// TIA Portal V20 export
FUNCTION_BLOCK "FB_Motor"   // FB102, LAD
TITLE = Direct-on-line motor with running feedback and trip monitoring
{ S7_Optimized_Access := 'TRUE' }
AUTHOR : Demo
VERSION : 0.2
// LAD version. Same interface as scl/14_FB_Motor.scl.
// stored: AutoNumber false, SetENOAutomatically false
   VAR_INPUT
      Run : Bool;   // Request: run the motor
      Permit : Bool := true;   // Interlock: motor may only run when TRUE
      RunFb : Bool;   // Running feedback (contactor auxiliary contact)
      Trip : Bool;   // Motor protection breaker tripped
      FeedbackTime : Time := T#5S;   // Max time from command to feedback
   END_VAR
   VAR_OUTPUT
      Out : Bool;   // Run command to the contactor
      Running : Bool;   // Motor confirmed running
      FaultTrip : Bool;   // Motor protection tripped
      FaultNoFeedback : Bool;   // Command on, but no running feedback within FeedbackTime
   END_VAR
   VAR
      tFb : TON_TIME;   // Feedback monitoring time
   END_VAR
BEGIN

REGION Network 1: Motor protection tripped
   // The motor protection breaker reports a trip.
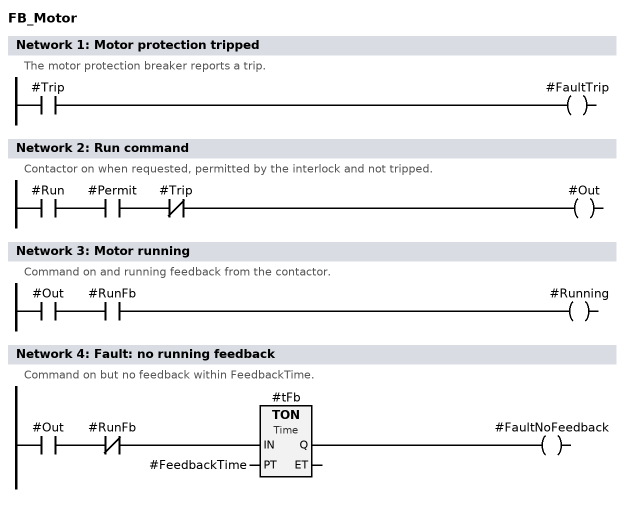
   RUNG wire#powerrail
      Contact( #Trip )
      Coil( #FaultTrip )
   END_RUNG
   // the same network as SCL:
   #FaultTrip := #Trip;
END_REGION

REGION Network 2: Run command
   // Contactor on when requested, permitted by the interlock and not tripped.
   RUNG wire#powerrail
      Contact( #Run )
      Contact( #Permit )
      I_Contact( #Trip )
      Coil( #Out )
   END_RUNG
   // the same network as SCL:
   #Out := #Run AND #Permit AND NOT #Trip;
END_REGION

REGION Network 3: Motor running
   // Command on and running feedback from the contactor.
   RUNG wire#powerrail
      Contact( #Out )
      Contact( #RunFb )
      Coil( #Running )
   END_RUNG
   // the same network as SCL:
   #Running := #Out AND #RunFb;
END_REGION

REGION Network 4: Fault: no running feedback
   // Command on but no feedback within FeedbackTime.
   RUNG wire#powerrail
      Contact( #Out )
      I_Contact( #RunFb )
      { S7_Templates := "time_type := Time" } #tFb.TON(pt := #FeedbackTime, et =>)
      Coil( #FaultNoFeedback )
   END_RUNG
   // the same network as SCL:
   #tFb(IN := #Out AND NOT #RunFb, PT := #FeedbackTime);   // TON
   #FaultNoFeedback := #tFb.Q;
END_REGION
END_FUNCTION_BLOCK
